      R_g[4,13] := -0.60548115;
      R_g[4,14] := 0.05480947;
      R_g[4,15] := 0.26145911;
      R_g[5,0] := 0.09851117;
      R_g[5,1] := 0.05978253;
      R_g[5,2] := -0.22380240;
      R_g[5,3] := 0.06287329;
      R_g[5,4] := 0.29527849;
      R_g[5,5] := -6.41728449;
      R_g[5,6] := -0.01966351;
      R_g[5,7] := 0.08289347;
      R_g[5,8] := 0.23354176;
      R_g[5,9] := 0.46406376;
      R_g[5,10] := -0.51907963;
      R_g[5,11] := -0.39992994;
      R_g[5,12] := 0.30295575;
      R_g[5,13] := 0.06150499;
      R_g[5,14] := -1.05495238;
      R_g[5,15] := -0.08431676;
      R_g[6,0] := -0.10256406;
      R_g[6,1] := 0.05051776;
      R_g[6,2] := 0.03060270;
      R_g[6,3] := 0.06608646;
      R_g[6,4] := -0.05028161;
      R_g[6,5] := -0.10387064;
      R_g[6,6] := -3.13754034;
      R_g[6,7] := -0.15655413;
      R_g[6,8] := 0.03909466;
      R_g[6,9] := -0.03506904;
      R_g[6,10] := 0.00484420;
      R_g[6,11] := -0.19064091;
      R_g[6,12] := 0.33072296;
      R_g[6,13] := -0.06755624;
      R_g[6,14] := -0.15698138;
      R_g[6,15] := -0.32207114;
      R_g[7,0] := 0.07863971;
      R_g[7,1] := -0.18754824;
      R_g[7,2] := -0.25378117;
      R_g[7,3] := -0.08824939;
      R_g[7,4] := -0.12941159;
      R_g[7,5] := 0.28854120;
      R_g[7,6] := 0.11216059;
      R_g[7,7] := -3.13675189;
      R_g[7,8] := -0.08472223;
      R_g[7,9] := 0.00790842;
      R_g[7,10] := -0.11386479;
      R_g[7,11] := -0.05684523;
      R_g[7,12] := 0.11065851;
      R_g[7,13] := -0.07569506;
      R_g[7,14] := 0.42330170;
      R_g[7,15] := -0.13425517;
      R_g[8,0] := 0.08961181;
      R_g[8,1] := 0.46519473;
      R_g[8,2] := -0.36562315;
      R_g[8,3] := 0.21113521;
      R_g[8,4] := -0.00757714;
      R_g[8,5] := -0.26392862;
      R_g[8,6] := 0.16387519;
      R_g[8,7] := -0.40587020;
      R_g[8,8] := -2.93437910;
      R_g[8,9] := 0.08376594;
      R_g[8,10] := -0.29606521;
      R_g[8,11] := 0.01828978;
      R_g[8,12] := 0.25248727;
      R_g[8,13] := -0.31344622;
      R_g[8,14] := -0.01567479;
      R_g[8,15] := 0.05443858;
      R_g[9,0] := -0.15096518;
      R_g[9,1] := -0.29858693;
      R_g[9,2] := 0.19766536;
      R_g[9,3] := -0.11255255;
      R_g[9,4] := -0.12072609;
      R_g[9,5] := 0.33710203;
      R_g[9,6] := 0.20158577;
      R_g[9,7] := -0.11389785;
      R_g[9,8] := -0.08645659;
      R_g[9,9] := -4.49089098;
      R_g[9,10] := 0.03153508;
      R_g[9,11] := 0.17591746;
      R_g[9,12] := -0.00816477;
      R_g[9,13] := -0.09244221;
      R_g[9,14] := -0.17023425;
      R_g[9,15] := 0.42906460;
      R_g[10,0] := -0.38857159;
      R_g[10,1] := 0.06436870;
      R_g[10,2] := -0.15642487;
      R_g[10,3] := -0.10405581;
      R_g[10,4] := 0.13234176;
      R_g[10,5] := 0.13661587;
      R_g[10,6] := 0.04957649;
      R_g[10,7] := 0.06489220;
      R_g[10,8] := 0.14693451;
      R_g[10,9] := -0.01300282;
      R_g[10,10] := -1.92830074;
      R_g[10,11] := 0.30045882;
      R_g[10,12] := 0.27313772;
      R_g[10,13] := 0.02955168;
      R_g[10,14] := -0.07842075;
      R_g[10,15] := 0.05753986;
      R_g[11,0] := -0.20971520;
      R_g[11,1] := 0.73070955;
      R_g[11,2] := -0.50315803;
      R_g[11,3] := 0.20500100;
      R_g[11,4] := -0.01089373;
      R_g[11,5] := 0.16404997;
      R_g[11,6] := 0.18906942;
      R_g[11,7] := 0.03491729;
      R_g[11,8] := -0.01610962;
      R_g[11,9] := 0.28074664;
      R_g[11,10] := 0.02013272;
      R_g[11,11] := -4.20378399;
      R_g[11,12] := 0.29341829;
      R_g[11,13] := 0.14369549;
      R_g[11,14] := -0.41985002;
      R_g[11,15] := 0.05762960;
      R_g[12,0] := -0.03705381;
      R_g[12,1] := -0.31124875;
      R_g[12,2] := 0.63473892;
      R_g[12,3] := 0.08633271;
      R_g[12,4] := -0.17926040;
      R_g[12,5] := 0.31777403;
      R_g[12,6] := -0.19864559;
      R_g[12,7] := -0.19772081;
      R_g[12,8] := 0.14220612;
      R_g[12,9] := -0.26425454;
      R_g[12,10] := 0.07095157;
      R_g[12,11] := 0.51232660;
      R_g[12,12] := -3.63068986;
      R_g[12,13] := -0.11757993;
      R_g[12,14] := 0.29906455;
      R_g[12,15] := -0.02980175;
      R_g[13,0] := 0.00863379;
      R_g[13,1] := 0.03295338;
      R_g[13,2] := -0.30022353;
      R_g[13,3] := 0.10327565;
      R_g[13,4] := -0.11605947;
      R_g[13,5] := 0.03122700;
      R_g[13,6] := 0.62577409;
      R_g[13,7] := 0.43430662;
      R_g[13,8] := 0.12523383;
      R_g[13,9] := 0.15241615;
      R_g[13,10] := -0.23994876;
      R_g[13,11] := -0.02434340;
      R_g[13,12] := 0.07577311;
      R_g[13,13] := -2.64277625;
      R_g[13,14] := -0.73717487;
      R_g[13,15] := -0.08735505;
      R_g[14,0] := -0.17141399;
      R_g[14,1] := 0.22617134;
      R_g[14,2] := -0.33173594;
      R_g[14,3] := 0.08776930;
      R_g[14,4] := 0.16216391;
      R_g[14,5] := 0.21827051;
      R_g[14,6] := 0.04451356;
      R_g[14,7] := 0.03265934;
      R_g[14,8] := -0.13619301;
      R_g[14,9] := 0.18478145;
      R_g[14,10] := -0.01089340;
      R_g[14,11] := -0.23413138;
      R_g[14,12] := 0.11226793;
      R_g[14,13] := 0.22237383;
      R_g[14,14] := -2.02859998;
      R_g[14,15] := -0.01800863;
      R_g[15,0] := 0.38834834;
      R_g[15,1] := -0.12119644;
      R_g[15,2] := -0.47133920;
      R_g[15,3] := 0.02589257;
      R_g[15,4] := -0.12965994;
      R_g[15,5] := -0.28714219;
      R_g[15,6] := 0.64088225;
      R_g[15,7] := 0.46508178;
      R_g[15,8] := -0.13015133;
      R_g[15,9] := 0.12145713;
      R_g[15,10] := 0.38442156;
      R_g[15,11] := -0.51173025;
      R_g[15,12] := -0.03178278;
      R_g[15,13] := -0.20804311;
      R_g[15,14] := 0.62473375;
      R_g[15,15] := -3.37922931;
      R_o[0,0] := -0.14847298;
      R_o[0,1] := -0.74705315;
      R_o[0,2] := 0.33793101;
      R_o[0,3] := 0.48812762;
      R_o[0,4] := -0.54246205;
      R_o[0,5] := 0.23658827;
      R_o[0,6] := 0.36877328;
      R_o[0,7] := -0.04479291;
      R_o[0,8] := 0.04525228;
      R_o[0,9] := -0.06947453;
      R_o[0,10] := -0.29408231;
      R_o[0,11] := -0.66140705;
      R_o[0,12] := -0.09016941;
      R_o[0,13] := -0.24453236;
      R_o[0,14] := 0.41733006;
      R_o[0,15] := 0.11528081;
      R_o[1,0] := -0.22536251;
      R_o[1,1] := -2.68759799;
      R_o[1,2] := 0.78251946;
      R_o[1,3] := 0.33114451;
      R_o[1,4] := -0.64871913;
      R_o[1,5] := -0.17744641;
      R_o[1,6] := -0.60721731;
      R_o[1,7] := -0.99844450;
      R_o[1,8] := 0.69376296;
      R_o[1,9] := -0.04945409;
      R_o[1,10] := 0.13805217;
      R_o[1,11] := 0.26013106;
      R_o[1,12] := -0.59883046;
      R_o[1,13] := -1.64951229;
      R_o[1,14] := -0.06540374;
      R_o[1,15] := -0.68399805;
      R_o[2,0] := 0.14265053;
      R_o[2,1] := -0.76361215;
      R_o[2,2] := 0.65221846;
      R_o[2,3] := -0.01308598;
      R_o[2,4] := -0.39565721;
      R_o[2,5] := -0.12863852;
      R_o[2,6] := 0.11177828;
      R_o[2,7] := -0.19651836;
      R_o[2,8] := 0.44556800;
      R_o[2,9] := -0.31979421;
      R_o[2,10] := 0.10245735;
      R_o[2,11] := -0.39614707;
      R_o[2,12] := -0.11074828;
      R_o[2,13] := -0.79570240;
      R_o[2,14] := 0.22064276;
      R_o[2,15] := 0.28490788;
      R_o[3,0] := 0.10347800;
      R_o[3,1] := -0.33515060;
      R_o[3,2] := 0.10071916;
      R_o[3,3] := 0.24764366;
      R_o[3,4] := -0.30636242;
      R_o[3,5] := -0.02347863;
      R_o[3,6] := 0.61475289;
      R_o[3,7] := 0.05460903;
      R_o[3,8] := -0.09153262;
      R_o[3,9] := -0.07667586;
      R_o[3,10] := 0.17097150;
      R_o[3,11] := -0.84717399;
      R_o[3,12] := 0.01488861;
      R_o[3,13] := 0.01246201;
      R_o[3,14] := 0.78524804;
      R_o[3,15] := -0.24291550;
      R_o[4,0] := 0.74034280;
      R_o[4,1] := -1.20240808;
      R_o[4,2] := -0.01728833;
      R_o[4,3] := -0.26750007;
      R_o[4,4] := 0.42328382;
      R_o[4,5] := -0.18842287;
      R_o[4,6] := -0.40243062;
      R_o[4,7] := 0.63144785;
      R_o[4,8] := -1.54348600;
      R_o[4,9] := 0.56258911;
      R_o[4,10] := -0.46023571;
      R_o[4,11] := -0.74631023;
      R_o[4,12] := 0.01794407;
      R_o[4,13] := 0.61756825;
      R_o[4,14] := -0.42400622;
      R_o[4,15] := -0.32165509;
      R_o[5,0] := -1.60871351;
      R_o[5,1] := -0.85439438;
      R_o[5,2] := 0.12367232;
      R_o[5,3] := 0.32163936;
      R_o[5,4] := -0.47827566;
      R_o[5,5] := 3.93251514;
      R_o[5,6] := -0.13689013;
      R_o[5,7] := 1.26777041;
      R_o[5,8] := -0.69722867;
      R_o[5,9] := -0.61384171;
      R_o[5,10] := 0.91998386;
      R_o[5,11] := -0.64498097;
      R_o[5,12] := -0.29473826;
      R_o[5,13] := -1.30750954;
      R_o[5,14] := 0.84536988;
      R_o[5,15] := 1.64059961;
      R_o[6,0] := 0.02413699;
      R_o[6,1] := -0.79112291;
      R_o[6,2] := -0.10358777;
      R_o[6,3] := -0.34534597;
      R_o[6,4] := 0.48224780;
      R_o[6,5] := -0.59422749;
      R_o[6,6] := 0.59001321;
      R_o[6,7] := 0.05578557;
      R_o[6,8] := -0.16264758;
      R_o[6,9] := -0.51271081;
      R_o[6,10] := 0.39541698;
      R_o[6,11] := -0.58911145;
      R_o[6,12] := -0.04537732;
      R_o[6,13] := 0.23783113;
      R_o[6,14] := 0.53961307;
      R_o[6,15] := 0.64036918;
      R_o[7,0] := 0.14012587;
      R_o[7,1] := -1.10767305;
      R_o[7,2] := 0.44994900;
      R_o[7,3] := 0.19807914;
      R_o[7,4] := -0.17633748;
      R_o[7,5] := -0.02624386;
      R_o[7,6] := 0.66549557;
      R_o[7,7] := 0.84196395;
      R_o[7,8] := 0.07700922;
      R_o[7,9] := 0.58576596;
      R_o[7,10] := 0.11728103;
      R_o[7,11] := -0.20590095;
      R_o[7,12] := -0.10266043;
      R_o[7,13] := 0.10980142;
      R_o[7,14] := 0.83650941;
      R_o[7,15] := 0.40667975;
      R_o[8,0] := 0.10407766;
      R_o[8,1] := -1.38828385;
      R_o[8,2] := 0.57484919;
      R_o[8,3] := -0.32096118;
      R_o[8,4] := -1.21653032;
      R_o[8,5] := -0.16445164;
      R_o[8,6] := 0.52185798;
      R_o[8,7] := 2.04115272;
      R_o[8,8] := -2.92285538;
      R_o[8,9] := -0.60037112;
      R_o[8,10] := -0.13611479;
      R_o[8,11] := -0.10244899;
      R_o[8,12] := -0.52569413;
      R_o[8,13] := -0.34149194;
      R_o[8,14] := 0.92290038;
      R_o[8,15] := -0.14947683;
      R_o[9,0] := 0.90203178;
      R_o[9,1] := -1.18227339;
      R_o[9,2] := 0.70378381;
      R_o[9,3] := -0.07063206;
      R_o[9,4] := -0.45001379;
      R_o[9,5] := 0.33594829;
      R_o[9,6] := 0.90896857;
      R_o[9,7] := -0.11313941;
      R_o[9,8] := 0.06154737;
      R_o[9,9] := -3.07011676;
      R_o[9,10] := 0.24497861;
      R_o[9,11] := -0.03553757;
      R_o[9,12] := -0.33283168;
      R_o[9,13] := 0.33938083;
      R_o[9,14] := 0.48779613;
      R_o[9,15] := 0.99066108;
      R_o[10,0] := 0.36748090;
      R_o[10,1] := -0.40652037;
      R_o[10,2] := 0.32123834;
      R_o[10,3] := 0.14693958;
      R_o[10,4] := -0.86366963;
      R_o[10,5] := 0.43876329;
      R_o[10,6] := -0.36798131;
      R_o[10,7] := -0.37096721;
      R_o[10,8] := 0.85877359;
      R_o[10,9] := -0.40861219;
      R_o[10,10] := 1.24025941;
      R_o[10,11] := -0.56068480;
      R_o[10,12] := -0.15937528;
      R_o[10,13] := -0.59108245;
      R_o[10,14] := 0.82221550;
      R_o[10,15] := 0.07025416;
      R_o[11,0] := -0.28333595;
      R_o[11,1] := -0.83661819;
      R_o[11,2] := 0.24413545;
      R_o[11,3] := 0.17671306;
      R_o[11,4] := -0.40138233;
      R_o[11,5] := 0.16249613;
      R_o[11,6] := 0.59071797;
      R_o[11,7] := 1.18243551;
      R_o[11,8] := -0.11446390;
      R_o[11,9] := -0.45934600;
      R_o[11,10] := 0.44795480;
      R_o[11,11] := 1.72437060;
      R_o[11,12] := -0.64456236;
      R_o[11,13] := -0.26468775;
      R_o[11,14] := 1.04931939;
      R_o[11,15] := 1.14608574;
      R_o[12,0] := 0.06811738;
      R_o[12,1] := -0.82940817;
      R_o[12,2] := 0.04298686;
      R_o[12,3] := 0.18846554;
      R_o[12,4] := -0.48880529;
      R_o[12,5] := 0.06246455;
      R_o[12,6] := 0.51301241;
      R_o[12,7] := 0.01585177;
      R_o[12,8] := -0.32864359;
      R_o[12,9] := -0.19140527;
      R_o[12,10] := 0.35500288;
      R_o[12,11] := -0.67324436;
      R_o[12,12] := -0.13675724;
      R_o[12,13] := 0.16862322;
      R_o[12,14] := 0.76524490;
      R_o[12,15] := 0.18042989;
      R_o[13,0] := 1.52919793;
      R_o[13,1] := -2.01665211;
      R_o[13,2] := 0.07069629;
      R_o[13,3] := 0.59324825;
      R_o[13,4] := -0.01248456;
      R_o[13,5] := 0.10036192;
      R_o[13,6] := 0.90690887;
      R_o[13,7] := 0.41812059;
      R_o[13,8] := -0.11101769;
      R_o[13,9] := -0.41462338;
      R_o[13,10] := 0.32745025;
      R_o[13,11] := 0.09499595;
      R_o[13,12] := -1.17409110;
      R_o[13,13] := 0.92265850;
      R_o[13,14] := 0.37988642;
      R_o[13,15] := 0.05125737;
      R_o[14,0] := 4.21519947;
      R_o[14,1] := -0.69102252;
      R_o[14,2] := 0.00603960;
      R_o[14,3] := -2.40963316;
      R_o[14,4] := -0.65538257;
      R_o[14,5] := -0.06152564;
      R_o[14,6] := -1.54533410;
      R_o[14,7] := -0.22543791;
      R_o[14,8] := 1.58575034;
      R_o[14,9] := -0.10917066;
      R_o[14,10] := 1.54773402;
      R_o[14,11] := -0.17321630;
      R_o[14,12] := -0.85895157;
      R_o[14,13] := -1.47213709;
      R_o[14,14] := 2.37665534;
      R_o[14,15] := -1.79636490;
      R_o[15,0] := 1.08996940;
      R_o[15,1] := -1.17211735;
      R_o[15,2] := 0.63166153;
      R_o[15,3] := 0.51676899;
      R_o[15,4] := -0.37341124;
      R_o[15,5] := 0.60133386;
      R_o[15,6] := 1.51174426;
      R_o[15,7] := 0.26480600;
      R_o[15,8] := 0.32437685;
      R_o[15,9] := -0.58537197;
      R_o[15,10] := -0.03915246;
      R_o[15,11] := -0.19543928;
      R_o[15,12] := -0.82763994;
      R_o[15,13] := 0.31273344;
      R_o[15,14] := 0.76913279;
      R_o[15,15] := 0.73493731;
      B_i[0] := -0.11525185;
      B_i[1] := -0.16767144;
      B_i[2] := -0.10675281;
      B_i[3] := 0.27595502;
      B_i[4] := 0.11127953;
      B_i[5] := -1.20700300;
      B_i[6] := -0.33555028;
      B_i[7] := -0.35219967;
      B_i[8] := -0.03516939;
      B_i[9] := -0.65995228;
      B_i[10] := 1.63097763;
      B_i[11] := -0.18333900;
      B_i[12] := 0.07472892;
      B_i[13] := 0.25719705;
      B_i[14] := -0.19151121;
      B_i[15] := -0.67595959;
      B_f[0] := 2.99556589;
      B_f[1] := -0.33741796;
      B_f[2] := 2.25157928;
      B_f[3] := 2.22067833;
      B_f[4] := -1.25157034;
      B_f[5] := 4.57832623;
      B_f[6] := 2.17673969;
      B_f[7] := 2.24434114;
      B_f[8] := 1.86623359;
      B_f[9] := 3.73503351;
      B_f[10] := 3.46735334;
      B_f[11] := 3.06714749;
      B_f[12] := 1.44914722;
      B_f[13] := 2.44668055;
      B_f[14] := 2.28946495;
      B_f[15] := 2.63645196;
      B_g[0] := 0.30800974;
      B_g[1] := -0.94244742;
      B_g[2] := 1.18943143;
      B_g[3] := 0.52035034;
      B_g[4] := 0.43232769;
      B_g[5] := 0.29648286;
      B_g[6] := 0.28049469;
      B_g[7] := 0.41938087;
      B_g[8] := -0.22911732;
      B_g[9] := -0.60563159;
      B_g[10] := 0.10972761;
      B_g[11] := 0.58977121;
      B_g[12] := -1.13596332;
      B_g[13] := 0.01335022;
      B_g[14] := 0.45130345;
      B_g[15] := 0.21969341;
      B_o[0] := 2.33575392;
      B_o[1] := 3.88747501;
      B_o[2] := 2.62646675;
      B_o[3] := 2.15524054;
      B_o[4] := 2.64990568;
      B_o[5] := 4.28425980;
      B_o[6] := 4.14953995;
      B_o[7] := 3.20074534;
      B_o[8] := 5.45463037;
      B_o[9] := 3.35326171;
      B_o[10] := 3.32303858;
      B_o[11] := 2.97783637;
      B_o[12] := 1.72812903;
      B_o[13] := 3.91121578;
      B_o[14] := 3.44036007;
      B_o[15] := 2.92046738;
      FC_W[0,0] := 0.76691687;
      FC_W[0,1] := 1.54350853;
      FC_W[0,2] := -0.20844251;
      FC_W[0,3] := 0.38317627;
      FC_W[0,4] := 0.75830436;
      FC_W[0,5] := 1.10985661;
      FC_W[0,6] := -0.95953107;
      FC_W[0,7] := 1.22366381;
      FC_W[0,8] := -0.21534167;
      FC_W[0,9] := -3.00756168;
      FC_W[0,10] := -0.08471649;
      FC_W[0,11] := 0.18020944;
      FC_W[0,12] := 0.58890468;
      FC_W[0,13] := -0.00262935;
      FC_W[0,14] := -0.60585809;
      FC_W[0,15] := 1.84203935;
      FC_W[1,0] := -0.84876847;
      FC_W[1,1] := -0.92502189;
      FC_W[1,2] := 0.94456464;
      FC_W[1,3] := -1.08595753;
      FC_W[1,4] := -0.52532524;
      FC_W[1,5] := 1.28364027;
      FC_W[1,6] := -2.58125854;
      FC_W[1,7] := -2.11014962;
      FC_W[1,8] := -0.25886634;
      FC_W[1,9] := -1.63888085;
      FC_W[1,10] := 0.76250589;
      FC_W[1,11] := 0.18522540;
      FC_W[1,12] := 1.45114386;
      FC_W[1,13] := -0.82991964;
      FC_W[1,14] := 1.54563367;
      FC_W[1,15] := -2.18503237;
      FC_W[2,0] := 0.74759591;
      FC_W[2,1] := 1.50420153;
      FC_W[2,2] := -0.13120306;
      FC_W[2,3] := 0.36578178;
      FC_W[2,4] := 0.76308554;
      FC_W[2,5] := 1.20159137;
      FC_W[2,6] := -1.16288304;
      FC_W[2,7] := 1.29092896;
      FC_W[2,8] := -0.21234436;
      FC_W[2,9] := -3.14010167;
      FC_W[2,10] := -0.10876910;
      FC_W[2,11] := 0.17469521;
      FC_W[2,12] := 0.70108241;
      FC_W[2,13] := 0.01334399;
      FC_W[2,14] := -0.75008494;
      FC_W[2,15] := 1.86712611;
      FC_W[3,0] := -0.45152566;
      FC_W[3,1] := 0.26790577;
      FC_W[3,2] := -0.35697538;
      FC_W[3,3] := -0.42768598;
      FC_W[3,4] := -0.15793064;
      FC_W[3,5] := -0.39237142;
      FC_W[3,6] := 1.28472209;
      FC_W[3,7] := -0.39581349;
      FC_W[3,8] := -0.63240361;
      FC_W[3,9] := -1.88796830;
      FC_W[3,10] := 0.01953238;
      FC_W[3,11] := 0.60719258;
      FC_W[3,12] := -0.00418234;
      FC_W[3,13] := 1.14158618;
      FC_W[3,14] := -0.57113940;
      FC_W[3,15] := -0.25580737;
      FC_W[4,0] := 1.29344773;
      FC_W[4,1] := -0.10325426;
      FC_W[4,2] := 0.57505780;
      FC_W[4,3] := -1.99647307;
      FC_W[4,4] := -0.48097378;
      FC_W[4,5] := -0.87535793;
      FC_W[4,6] := 0.76299852;
      FC_W[4,7] := -0.31900346;
      FC_W[4,8] := 0.43593013;
      FC_W[4,9] := 0.34549168;
      FC_W[4,10] := 0.01366996;
      FC_W[4,11] := 1.01956534;
      FC_W[4,12] := -0.61152214;
      FC_W[4,13] := -1.56243253;
      FC_W[4,14] := -1.10839498;
      FC_W[4,15] := 1.56659317;
      FC_W[5,0] := 0.41176695;
      FC_W[5,1] := -1.24408734;
      FC_W[5,2] := 0.48085922;
      FC_W[5,3] := 1.40249288;
      FC_W[5,4] := -0.05570108;
      FC_W[5,5] := -6.80598259;
      FC_W[5,6] := -0.69677407;
      FC_W[5,7] := 0.74036807;
      FC_W[5,8] := 1.61717665;
      FC_W[5,9] := -0.05372217;
      FC_W[5,10] := -1.22660577;
      FC_W[5,11] := 0.25594920;
      FC_W[5,12] := 0.23262075;
      FC_W[5,13] := -0.50597012;
      FC_W[5,14] := 0.23332803;
      FC_W[5,15] := -0.61406231;
      FC_W[6,0] := 0.61248779;
      FC_W[6,1] := 1.53917146;
      FC_W[6,2] := -0.01028113;
      FC_W[6,3] := 0.66907030;
      FC_W[6,4] := -0.14260414;
      FC_W[6,5] := -1.26385117;
      FC_W[6,6] := -0.33451670;
      FC_W[6,7] := 0.33876544;
      FC_W[6,8] := 0.47751576;
      FC_W[6,9] := 0.96330714;
      FC_W[6,10] := -0.17724371;
      FC_W[6,11] := 2.24375200;
      FC_W[6,12] := -0.40486264;
      FC_W[6,13] := 0.65613246;
      FC_W[6,14] := -0.44845906;
      FC_W[6,15] := -0.68273169;
      FC_W[7,0] := -0.44028389;
      FC_W[7,1] := 0.29088175;
      FC_W[7,2] := -0.38207194;
      FC_W[7,3] := -0.41779745;
      FC_W[7,4] := -0.17482910;
      FC_W[7,5] := -0.42837557;
      FC_W[7,6] := 1.36843240;
      FC_W[7,7] := -0.39042190;
      FC_W[7,8] := -0.62430942;
      FC_W[7,9] := -1.80241871;
      FC_W[7,10] := 0.04712024;
      FC_W[7,11] := 0.60730672;
      FC_W[7,12] := -0.07031967;
      FC_W[7,13] := 1.14298403;
      FC_W[7,14] := -0.52446443;
      FC_W[7,15] := -0.25127152;
      FC_W[8,0] := -0.50533390;
      FC_W[8,1] := 0.30554622;
      FC_W[8,2] := -0.38464165;
      FC_W[8,3] := -0.48505715;
      FC_W[8,4] := -0.07984031;
      FC_W[8,5] := -0.35821158;
      FC_W[8,6] := 1.20251560;
      FC_W[8,7] := -0.44205466;
      FC_W[8,8] := -0.64952880;
      FC_W[8,9] := -2.03045917;
      FC_W[8,10] := 0.04362446;
      FC_W[8,11] := 0.59587187;
      FC_W[8,12] := 0.12079757;
      FC_W[8,13] := 1.11798072;
      FC_W[8,14] := -0.63356131;
      FC_W[8,15] := -0.29604205;
      FC_W[9,0] := -0.45088705;
      FC_W[9,1] := 0.27602863;
      FC_W[9,2] := -0.37352136;
      FC_W[9,3] := -0.41263905;
      FC_W[9,4] := -0.16068281;
      FC_W[9,5] := -0.40061781;
      FC_W[9,6] := 1.31766760;
      FC_W[9,7] := -0.38225642;
      FC_W[9,8] := -0.63187581;
      FC_W[9,9] := -1.85595226;
      FC_W[9,10] := 0.04726556;
      FC_W[9,11] := 0.59707093;
      FC_W[9,12] := -0.02673960;
      FC_W[9,13] := 1.14315939;
      FC_W[9,14] := -0.53523809;
      FC_W[9,15] := -0.25229296;
      FC_W[10,0] := -1.11255634;
      FC_W[10,1] := -1.10758793;
      FC_W[10,2] := -0.24714845;
      FC_W[10,3] := -0.59940976;
      FC_W[10,4] := -0.10819428;
      FC_W[10,5] := -1.58778656;
      FC_W[10,6] := 0.60180962;
      FC_W[10,7] := -0.69662166;
      FC_W[10,8] := -0.63675028;
      FC_W[10,9] := -3.21672893;
      FC_W[10,10] := 0.03261364;
      FC_W[10,11] := -1.07562602;
      FC_W[10,12] := 0.92825305;
      FC_W[10,13] := 0.36362201;
      FC_W[10,14] := 0.14236267;
      FC_W[10,15] := -0.23976374;
      FC_W[11,0] := -0.03737991;
      FC_W[11,1] := -0.06299526;
      FC_W[11,2] := 0.61952871;
      FC_W[11,3] := 0.19341917;
      FC_W[11,4] := -1.42015672;
      FC_W[11,5] := 0.08432721;
      FC_W[11,6] := 0.30952653;
      FC_W[11,7] := 0.81136137;
      FC_W[11,8] := -1.67836761;
      FC_W[11,9] := -0.01523663;
      FC_W[11,10] := -0.87199742;
      FC_W[11,11] := 0.11922295;
      FC_W[11,12] := 0.38131532;
      FC_W[11,13] := -0.28784695;
      FC_W[11,14] := -0.13377608;
      FC_W[11,15] := -0.11664936;
      FC_W[12,0] := -0.21013576;
      FC_W[12,1] := -0.25084072;
      FC_W[12,2] := 0.69950396;
      FC_W[12,3] := 0.10803718;
      FC_W[12,4] := -1.51941526;
      FC_W[12,5] := 0.05514818;
      FC_W[12,6] := -0.01964889;
      FC_W[12,7] := 1.25729561;
      FC_W[12,8] := -1.13359058;
      FC_W[12,9] := -0.04563072;
      FC_W[12,10] := -0.36160040;
      FC_W[12,11] := -0.04378428;
      FC_W[12,12] := 0.12715936;
      FC_W[12,13] := -0.02202382;
      FC_W[12,14] := -0.23011394;
      FC_W[12,15] := -0.30061662;
      FC_W[13,0] := 0.74089515;
      FC_W[13,1] := -0.07237465;
      FC_W[13,2] := 0.01080942;
      FC_W[13,3] := -0.13760488;
      FC_W[13,4] := -0.40318596;
      FC_W[13,5] := 0.09405857;
      FC_W[13,6] := -0.62446254;
      FC_W[13,7] := 0.10771502;
      FC_W[13,8] := -0.52130091;
      FC_W[13,9] := -0.55923247;
      FC_W[13,10] := 2.08023214;
      FC_W[13,11] := -0.26325747;
      FC_W[13,12] := -0.60065490;
      FC_W[13,13] := 0.73370737;
      FC_W[13,14] := 4.43074036;
      FC_W[13,15] := -1.03970754;
      FC_W[14,0] := -3.11080956;
      FC_W[14,1] := 1.52514708;
      FC_W[14,2] := -0.30008835;
      FC_W[14,3] := -3.75322127;
      FC_W[14,4] := 0.61758131;
      FC_W[14,5] := 0.79863137;
      FC_W[14,6] := 0.85665506;
      FC_W[14,7] := 2.64684296;
      FC_W[14,8] := 1.93208790;
      FC_W[14,9] := -0.02786120;
      FC_W[14,10] := -3.76214457;
      FC_W[14,11] := 2.24488688;
      FC_W[14,12] := 2.17172313;
      FC_W[14,13] := 0.52849472;
      FC_W[14,14] := 2.06621265;
      FC_W[14,15] := 0.21302631;
      FC_W[15,0] := 0.16616058;
      FC_W[15,1] := 0.10622021;
      FC_W[15,2] := 0.53326297;
      FC_W[15,3] := 0.31807119;
      FC_W[15,4] := -1.17440403;
      FC_W[15,5] := 0.08476182;
      FC_W[15,6] := 0.11705037;
      FC_W[15,7] := -0.01000034;
      FC_W[15,8] := -2.36726975;
      FC_W[15,9] := 0.03094000;
      FC_W[15,10] := -1.62616897;
      FC_W[15,11] := 0.33965093;
      FC_W[15,12] := 0.60757959;
      FC_W[15,13] := -0.14965913;
      FC_W[15,14] := -0.00611463;
      FC_W[15,15] := 0.40740597;
      FC_W[16,0] := -0.96380889;
      FC_W[16,1] := 1.08168781;
      FC_W[16,2] := 2.37668490;
      FC_W[16,3] := -1.05731308;
      FC_W[16,4] := 0.29249096;
      FC_W[16,5] := -0.36915782;
      FC_W[16,6] := -3.40412092;
      FC_W[16,7] := -3.52345991;
      FC_W[16,8] := -0.07057770;
      FC_W[16,9] := 0.63422161;
      FC_W[16,10] := -1.44417024;
      FC_W[16,11] := -0.88294816;
      FC_W[16,12] := 0.74554622;
      FC_W[16,13] := 4.62807751;
      FC_W[16,14] := 0.40313786;
      FC_W[16,15] := 3.93857050;
      FC_W[17,0] := -1.18036187;
      FC_W[17,1] := -0.28546566;
      FC_W[17,2] := 1.83997035;
      FC_W[17,3] := -0.86653274;
      FC_W[17,4] := -0.62797892;
      FC_W[17,5] := -0.24189699;
      FC_W[17,6] := -1.59377563;
      FC_W[17,7] := 3.17389417;
      FC_W[17,8] := 4.20314360;
      FC_W[17,9] := 0.37900031;
      FC_W[17,10] := 3.86766505;
      FC_W[17,11] := -2.21274209;
      FC_W[17,12] := -1.37958419;
      FC_W[17,13] := 1.73672819;
      FC_W[17,14] := -0.71695817;
      FC_W[17,15] := -1.04806626;
      FC_W[18,0] := 0.16363387;
      FC_W[18,1] := 2.46524715;
      FC_W[18,2] := -0.78923774;
      FC_W[18,3] := 0.87476426;
      FC_W[18,4] := -5.95409679;
      FC_W[18,5] := 0.88954771;
      FC_W[18,6] := 1.85371697;
      FC_W[18,7] := -0.90911502;
      FC_W[18,8] := 1.67899203;
      FC_W[18,9] := 0.08326869;
      FC_W[18,10] := -0.33310106;
      FC_W[18,11] := -1.37995827;
      FC_W[18,12] := 0.17668670;
      FC_W[18,13] := -1.74094355;
      FC_W[18,14] := -0.14677437;
      FC_W[18,15] := 0.79526556;
      FC_W[19,0] := -0.25457042;
      FC_W[19,1] := -0.94162971;
      FC_W[19,2] := 0.57019746;
      FC_W[19,3] := -0.06669754;
      FC_W[19,4] := -0.31895879;
      FC_W[19,5] := -0.11969372;
      FC_W[19,6] := -0.37630516;
      FC_W[19,7] := 1.84739316;
      FC_W[19,8] := -1.24445868;
      FC_W[19,9] := -0.09252350;
      FC_W[19,10] := -0.06256182;
      FC_W[19,11] := 0.33049041;
      FC_W[19,12] := -0.05521645;
      FC_W[19,13] := 0.08963338;
      FC_W[19,14] := -0.24520318;
      FC_W[19,15] := -0.76362497;
      FC_W[20,0] := -0.44794476;
      FC_W[20,1] := -2.14960837;
      FC_W[20,2] := 0.29591742;
      FC_W[20,3] := -0.17743635;
      FC_W[20,4] := -0.58367479;
      FC_W[20,5] := 0.58847088;
      FC_W[20,6] := 1.35463679;
      FC_W[20,7] := -0.16127646;
      FC_W[20,8] := -0.27197161;
      FC_W[20,9] := -0.63772136;
      FC_W[20,10] := 0.51769370;
      FC_W[20,11] := -1.32718563;
      FC_W[20,12] := 0.35489064;
      FC_W[20,13] := -0.78381717;
      FC_W[20,14] := 0.89823222;
      FC_W[20,15] := 1.42503154;
      FC_W[21,0] := -2.43106961;
      FC_W[21,1] := 1.03015459;
      FC_W[21,2] := -0.23634396;
      FC_W[21,3] := 1.30044115;
      FC_W[21,4] := 0.44065619;
      FC_W[21,5] := 0.70075428;
      FC_W[21,6] := -0.38531300;
      FC_W[21,7] := 0.12913185;
      FC_W[21,8] := -0.46658489;
      FC_W[21,9] := -0.65548015;
      FC_W[21,10] := 0.36299118;
      FC_W[21,11] := 1.43775284;
      FC_W[21,12] := -0.36456382;
      FC_W[21,13] := -0.45043552;
      FC_W[21,14] := -0.56249213;
      FC_W[21,15] := 1.26511896;
      FC_W[22,0] := 0.22401933;
      FC_W[22,1] := -1.52788472;
      FC_W[22,2] := 2.09116197;
      FC_W[22,3] := 0.56461936;
      FC_W[22,4] := -0.46243390;
      FC_W[22,5] := 0.73684770;
      FC_W[22,6] := 0.19164361;
      FC_W[22,7] := 0.06346934;
      FC_W[22,8] := 0.54199892;
      FC_W[22,9] := -1.03965259;
      FC_W[22,10] := -0.24938214;
      FC_W[22,11] := 2.15651417;
      FC_W[22,12] := -1.79916179;
      FC_W[22,13] := -0.21550527;
      FC_W[22,14] := 0.60506076;
      FC_W[22,15] := 0.58267546;
      FC_W[23,0] := 0.93549359;
      FC_W[23,1] := -0.40594038;
      FC_W[23,2] := -0.16483921;
      FC_W[23,3] := 0.02804452;
      FC_W[23,4] := -0.54419273;
      FC_W[23,5] := -0.10059550;
      FC_W[23,6] := 0.57842124;
      FC_W[23,7] := -0.12527937;
      FC_W[23,8] := -0.78040689;
      FC_W[23,9] := -0.61837119;
      FC_W[23,10] := 1.44107115;
      FC_W[23,11] := -0.16925113;
      FC_W[23,12] := -0.83583456;
      FC_W[23,13] := 1.60294521;
      FC_W[23,14] := 4.23907661;
      FC_W[23,15] := -1.32083130;
      FC_W[24,0] := 0.18377206;
      FC_W[24,1] := -1.39490736;
      FC_W[24,2] := 1.99884033;
      FC_W[24,3] := 0.55039299;
      FC_W[24,4] := -0.58098501;
      FC_W[24,5] := 0.63703549;
      FC_W[24,6] := 0.29183668;
      FC_W[24,7] := 0.03679674;
      FC_W[24,8] := 0.54975742;
      FC_W[24,9] := -0.83437216;
      FC_W[24,10] := -0.22163391;
      FC_W[24,11] := 2.07142234;
      FC_W[24,12] := -2.01642585;
      FC_W[24,13] := -0.23686101;
      FC_W[24,14] := 0.70799166;
      FC_W[24,15] := 0.58019441;
      FC_W[25,0] := 0.18751292;
      FC_W[25,1] := -1.40110946;
      FC_W[25,2] := 2.01208258;
      FC_W[25,3] := 0.55488765;
      FC_W[25,4] := -0.58586031;
      FC_W[25,5] := 0.63924384;
      FC_W[25,6] := 0.29609177;
      FC_W[25,7] := 0.03836685;
      FC_W[25,8] := 0.55524427;
      FC_W[25,9] := -0.83095372;
      FC_W[25,10] := -0.22373353;
      FC_W[25,11] := 2.08144498;
      FC_W[25,12] := -2.02489543;
      FC_W[25,13] := -0.23646893;
      FC_W[25,14] := 0.70846170;
      FC_W[25,15] := 0.58629918;
      FC_W[26,0] := 1.66300058;
      FC_W[26,1] := -1.82226586;
      FC_W[26,2] := 1.66785717;
      FC_W[26,3] := -0.62902045;
      FC_W[26,4] := 0.32130203;
      FC_W[26,5] := -0.16516249;
      FC_W[26,6] := -0.31834188;
      FC_W[26,7] := -0.01305876;
      FC_W[26,8] := 0.24688217;
      FC_W[26,9] := -0.64328623;
      FC_W[26,10] := -0.01610377;
      FC_W[26,11] := 1.13409078;
      FC_W[26,12] := -0.77092558;
      FC_W[26,13] := 0.59138787;
      FC_W[26,14] := 1.18435347;
      FC_W[26,15] := -0.78926718;
      FC_W[27,0] := -2.89214182;
      FC_W[27,1] := 1.40610170;
      FC_W[27,2] := -0.86616915;
      FC_W[27,3] := 0.77281964;
      FC_W[27,4] := 0.79401380;
      FC_W[27,5] := 0.34485626;
      FC_W[27,6] := -0.39616618;
      FC_W[27,7] := -0.09319982;
      FC_W[27,8] := -0.91662061;
      FC_W[27,9] := -0.42657280;
      FC_W[27,10] := 0.81243485;
      FC_W[27,11] := 0.88650566;
      FC_W[27,12] := -0.40733227;
      FC_W[27,13] := -0.55559754;
      FC_W[27,14] := -0.23531459;
      FC_W[27,15] := 1.34971523;
      FC_W[28,0] := 1.56295800;
      FC_W[28,1] := 1.42122293;
      FC_W[28,2] := 0.00074465;
      FC_W[28,3] := -2.07726741;
      FC_W[28,4] := 0.43710080;
      FC_W[28,5] := -1.41943741;
      FC_W[28,6] := -0.53313965;
      FC_W[28,7] := -0.04702906;
      FC_W[28,8] := -0.36702093;
      FC_W[28,9] := 0.37743872;
      FC_W[28,10] := 0.59604365;
      FC_W[28,11] := 2.10622239;
      FC_W[28,12] := 0.02389226;
      FC_W[28,13] := -0.84609389;
      FC_W[28,14] := -0.47065067;
      FC_W[28,15] := 0.46141356;
      FC_W[29,0] := 0.18336056;
      FC_W[29,1] := 1.35958064;
      FC_W[29,2] := -1.92125678;
      FC_W[29,3] := -0.44665357;
      FC_W[29,4] := 0.67866659;
      FC_W[29,5] := -1.27040529;
      FC_W[29,6] := 0.34309217;
      FC_W[29,7] := 0.30406588;
      FC_W[29,8] := -0.28503451;
      FC_W[29,9] := 2.14690542;
      FC_W[29,10] := -0.13428468;
      FC_W[29,11] := -2.26440001;
      FC_W[29,12] := 0.57903779;
      FC_W[29,13] := 0.48088390;
      FC_W[29,14] := -0.51877141;
      FC_W[29,15] := -0.67464572;
      FC_W[30,0] := 0.22795415;
      FC_W[30,1] := -1.53159809;
      FC_W[30,2] := 2.09372473;
      FC_W[30,3] := 0.56482655;
      FC_W[30,4] := -0.46061462;
      FC_W[30,5] := 0.73824251;
      FC_W[30,6] := 0.18884818;
      FC_W[30,7] := 0.06514335;
      FC_W[30,8] := 0.54162019;
      FC_W[30,9] := -1.04339278;
      FC_W[30,10] := -0.25149027;
      FC_W[30,11] := 2.15671182;
      FC_W[30,12] := -1.79456043;
      FC_W[30,13] := -0.21399722;
      FC_W[30,14] := 0.60102427;
      FC_W[30,15] := 0.58390999;
      FC_W[31,0] := 0.27823162;
      FC_W[31,1] := -1.58497131;
      FC_W[31,2] := 2.12941575;
      FC_W[31,3] := 0.57324249;
      FC_W[31,4] := -0.40936530;
      FC_W[31,5] := 0.77423245;
      FC_W[31,6] := 0.17383640;
      FC_W[31,7] := 0.10636473;
      FC_W[31,8] := 0.55564606;
      FC_W[31,9] := -1.07348740;
      FC_W[31,10] := -0.28553542;
      FC_W[31,11] := 2.19243288;
      FC_W[31,12] := -1.70922673;
      FC_W[31,13] := -0.19247352;
      FC_W[31,14] := 0.52959895;
      FC_W[31,15] := 0.59279895;
      FC_W[32,0] := 0.04953038;
      FC_W[32,1] := -1.41549408;
      FC_W[32,2] := 2.01636505;
      FC_W[32,3] := 0.50114906;
      FC_W[32,4] := -0.46179849;
      FC_W[32,5] := 0.74877977;
      FC_W[32,6] := 0.13434805;
      FC_W[32,7] := -0.03319941;
      FC_W[32,8] := 0.45586070;
      FC_W[32,9] := -1.14118552;
      FC_W[32,10] := -0.13540792;
      FC_W[32,11] := 2.23494720;
      FC_W[32,12] := -1.73130178;
      FC_W[32,13] := -0.31032586;
      FC_W[32,14] := 0.63603759;
      FC_W[32,15] := 0.65046942;
      FC_W[33,0] := -0.00627907;
      FC_W[33,1] := -1.49908721;
      FC_W[33,2] := 2.07251692;
      FC_W[33,3] := 0.47237280;
      FC_W[33,4] := -0.28603134;
      FC_W[33,5] := 0.86122340;
      FC_W[33,6] := -0.05305826;
      FC_W[33,7] := -0.05858019;
      FC_W[33,8] := 0.40629035;
      FC_W[33,9] := -1.41835237;
      FC_W[33,10] := -0.12844640;
      FC_W[33,11] := 2.38462377;
      FC_W[33,12] := -1.41297781;
      FC_W[33,13] := -0.36302483;
      FC_W[33,14] := 0.44525054;
      FC_W[33,15] := 0.69628060;
      FC_W[34,0] := 0.08176677;
      FC_W[34,1] := -1.52486050;
      FC_W[34,2] := 2.10055542;
      FC_W[34,3] := 0.50965518;
      FC_W[34,4] := -0.35586321;
      FC_W[34,5] := 0.87471449;
      FC_W[34,6] := 0.00432379;
      FC_W[34,7] := -0.01442015;
      FC_W[34,8] := 0.46000737;
      FC_W[34,9] := -1.38360655;
      FC_W[34,10] := -0.18607068;
      FC_W[34,11] := 2.33854008;
      FC_W[34,12] := -1.44122565;
      FC_W[34,13] := -0.33802593;
      FC_W[34,14] := 0.43794119;
      FC_W[34,15] := 0.68164617;
      FC_W[35,0] := 0.00513690;
      FC_W[35,1] := -1.32884324;
      FC_W[35,2] := 1.90931404;
      FC_W[35,3] := 0.49852094;
      FC_W[35,4] := -0.56343287;
      FC_W[35,5] := 0.67876500;
      FC_W[35,6] := 0.23343433;
      FC_W[35,7] := -0.06241892;
      FC_W[35,8] := 0.42093012;
      FC_W[35,9] := -1.01738036;
      FC_W[35,10] := -0.03109938;
      FC_W[35,11] := 2.15396738;
      FC_W[35,12] := -1.84033465;
      FC_W[35,13] := -0.29486498;
      FC_W[35,14] := 0.83844137;
      FC_W[35,15] := 0.63658357;
      FC_W[36,0] := -1.56804621;
      FC_W[36,1] := 1.12077355;
      FC_W[36,2] := 0.21489759;
      FC_W[36,3] := -0.85609603;
      FC_W[36,4] := 0.41929087;
      FC_W[36,5] := -0.72125524;
      FC_W[36,6] := -0.20861968;
      FC_W[36,7] := -0.47542524;
      FC_W[36,8] := 0.05816720;
      FC_W[36,9] := 0.88530207;
      FC_W[36,10] := -1.33813703;
      FC_W[36,11] := -1.43648410;
      FC_W[36,12] := -6.04789782;
      FC_W[36,13] := -0.41200089;
      FC_W[36,14] := 0.47274289;
      FC_W[36,15] := -0.30960068;
      FC_W[37,0] := -0.01744911;
      FC_W[37,1] := -1.28811061;
      FC_W[37,2] := 1.87406683;
      FC_W[37,3] := 0.49300796;
      FC_W[37,4] := -0.57639700;
      FC_W[37,5] := 0.65250272;
      FC_W[37,6] := 0.24592924;
      FC_W[37,7] := -0.07283052;
      FC_W[37,8] := 0.40504485;
      FC_W[37,9] := -0.97370982;
      FC_W[37,10] := -0.00745488;
      FC_W[37,11] := 2.12590337;
      FC_W[37,12] := -1.89184034;
      FC_W[37,13] := -0.28358787;
      FC_W[37,14] := 0.89717782;
      FC_W[37,15] := 0.61702895;
      FC_W[38,0] := -0.28529665;
      FC_W[38,1] := -2.81238103;
      FC_W[38,2] := -3.51768899;
      FC_W[38,3] := 0.40109450;
      FC_W[38,4] := -0.98214322;
      FC_W[38,5] := 0.33394021;
      FC_W[38,6] := -3.25278091;
      FC_W[38,7] := -1.33008122;
      FC_W[38,8] := 0.27982229;
      FC_W[38,9] := -1.03831351;
      FC_W[38,10] := 0.04537877;
      FC_W[38,11] := 2.10162973;
      FC_W[38,12] := -1.06387031;
      FC_W[38,13] := 1.87411618;
      FC_W[38,14] := -0.54168665;
      FC_W[38,15] := 1.84349597;
      FC_W[39,0] := -1.92901528;
      FC_W[39,1] := -0.78533107;
      FC_W[39,2] := -2.23502517;
      FC_W[39,3] := -1.94082272;
      FC_W[39,4] := -0.12267892;
      FC_W[39,5] := 0.66615528;
      FC_W[39,6] := -1.05431843;
      FC_W[39,7] := 1.03078413;
      FC_W[39,8] := 1.43677998;
      FC_W[39,9] := -0.67489189;
      FC_W[39,10] := -2.09733391;
      FC_W[39,11] := 2.61480737;
      FC_W[39,12] := 0.58990037;
      FC_W[39,13] := 1.10489023;
      FC_W[39,14] := 0.74517161;
      FC_W[39,15] := 0.87154233;
      FC_B[0] := -0.33364403;
      FC_B[1] := -0.07630836;
      FC_B[2] := -0.34703955;
      FC_B[3] := 0.05934331;
      FC_B[4] := -0.66695452;
      FC_B[5] := -0.13967955;
      FC_B[6] := 0.48994508;
      FC_B[7] := 0.06493863;
      FC_B[8] := 0.09218118;
      FC_B[9] := 0.06467691;
      FC_B[10] := -0.19661079;
      FC_B[11] := -0.49837264;
      FC_B[12] := -0.48156646;
      FC_B[13] := -0.83966696;
      FC_B[14] := 0.72801244;
      FC_B[15] := -0.50594783;
      FC_B[16] := 0.14493598;
      FC_B[17] := 0.02873158;
      FC_B[18] := 1.81477070;
      FC_B[19] := -0.81444138;
      FC_B[20] := -0.82179058;
      FC_B[21] := 0.40513784;
      FC_B[22] := -1.70836389;
      FC_B[23] := -0.88778102;
      FC_B[24] := -1.65490472;
      FC_B[25] := -1.66285884;
      FC_B[26] := -1.66001046;
      FC_B[27] := 0.64861679;
      FC_B[28] := -0.22430785;
      FC_B[29] := 1.42981255;
      FC_B[30] := -1.70972085;
      FC_B[31] := -1.72291648;
      FC_B[32] := -1.65422285;
      FC_B[33] := -1.66723549;
      FC_B[34] := -1.67813110;
      FC_B[35] := -1.61601245;
      FC_B[36] := -0.68123728;
      FC_B[37] := -1.60075045;
      FC_B[38] := 0.83955693;
      FC_B[39] := 0.87614125;

END_DATA_BLOCK
